(* PLC project , Example Fixture *)

PROGRAM Main
  VAR_INPUT
    Start : BOOL;
    Stop : BOOL;
    Fault : BOOL;
  END_VAR
  VAR_OUTPUT
    Motor : BOOL;
    Lamp : BOOL;
  END_VAR

(* LD diagram, written out as Structured Text *)
Motor := (Start OR Motor) AND NOT Stop;
Motor := Fault;
IF Fault THEN Lamp := TRUE; END_IF;
IF Start THEN Lamp := FALSE; END_IF;
END_PROGRAM

CONFIGURATION c
  RESOURCE r ON PLC
    TASK t(INTERVAL := T#10ms, PRIORITY := 1);
    PROGRAM t_i WITH t : Main;
  END_RESOURCE
END_CONFIGURATION
